Fanuc KAREL source: KA00050.KL

PROGRAM KA00050
%NOLOCKGROUP
VAR
  SRC: POSITION
  DST: REAL
BEGIN
  DST = SRC
END KA00050
